DATA_BLOCK "FRK_Load_D008A"
{ S7_Optimized_Access := 'TRUE' }
VERSION : 0.1
UNLINKED
NON_RETAIN
VAR
    Bytes {ExternalAccessible := 'False'; ExternalVisible := 'False'; ExternalWritable := 'False'} : Array[0..8249] of Byte;
END_VAR
BEGIN
END_DATA_BLOCK
